(* CODESYS project EVs.export

Project tree, tasks and I/O mapping:
  visualisation EVs
*)

// /EVs
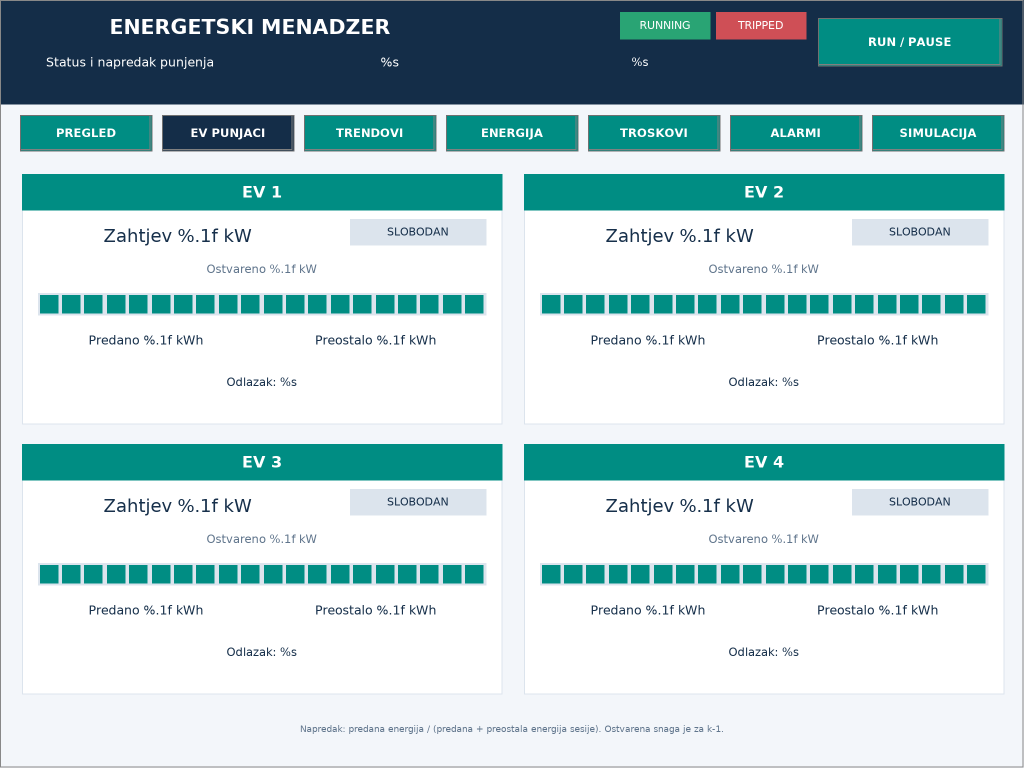
VISUALIZATION EVs  // 1024x768
    Rectangle (0,0 1024x768)
    Rectangle (0,0 1024x104)
    Rectangle (20,10 460x34), "ENERGETSKI MENADZER"
    Rectangle (20,48 220x28), "Status i napredak punjenja"
    Rectangle (260,49 260x26), "%s", text variable: Team_HMI.sDateTime
    Rectangle (530,49 220x26), "%s", text variable: Team_HMI.sPriceMode
    Button (818,18 184x48), "RUN / PAUSE"
        toggle SimCtrl.run
    Rectangle (620,12 90x27), "PAUSED", invisible if: SimCtrl.run
    Rectangle (620,12 90x27), "RUNNING", invisible if: NOT SimCtrl.run
    Rectangle (716,12 90x27), "TRIPPED", invisible if: NOT SimCtrl.tripped
    Button (20,115 132x36), "PREGLED"
        OnMouseClick:  Assign=Overview, Type=Assignment
    Button (162,115 132x36), "EV PUNJACI"
        OnMouseClick:  Assign=EVs, Type=Assignment
    Button (304,115 132x36), "TRENDOVI"
        OnMouseClick:  Assign=Trends, Type=Assignment
    Button (446,115 132x36), "ENERGIJA"
        OnMouseClick:  Assign=Energy, Type=Assignment
    Button (588,115 132x36), "TROSKOVI"
        OnMouseClick:  Assign=Costs, Type=Assignment
    Button (730,115 132x36), "ALARMI"
        OnMouseClick:  Assign=Alarms, Type=Assignment
    Button (872,115 132x36), "SIMULACIJA"
        OnMouseClick:  Assign=Controls, Type=Assignment
    Rectangle (22,174 480x250)
    Rectangle (22,174 480x36), "EV 1"
    Rectangle (350,219 136x26), "SPOJEN", invisible if: NOT Team_HMI.aEvConnected[0]
    Rectangle (350,219 136x26), "SLOBODAN", invisible if: Team_HMI.aEvConnected[0]
    Rectangle (38,218 280x36), "Zahtjev %.1f kW", text variable: Team_HMI.aEvReq[0]
    Rectangle (38,256 448x26), "Ostvareno %.1f kW", text variable: Team_HMI.aEvAct[0]
    Rectangle (38,293 448x22)
    Rectangle (40,295 18x18), invisible if: (100.0 * Team_HMI.aEvDelivered[0] / MAX(0.001, Team_HMI.aEvDelivered[0] + Team_HMI.aEvRemaining[0])) < 5.000
    Rectangle (62,295 18x18), invisible if: (100.0 * Team_HMI.aEvDelivered[0] / MAX(0.001, Team_HMI.aEvDelivered[0] + Team_HMI.aEvRemaining[0])) < 10.000
    Rectangle (84,295 18x18), invisible if: (100.0 * Team_HMI.aEvDelivered[0] / MAX(0.001, Team_HMI.aEvDelivered[0] + Team_HMI.aEvRemaining[0])) < 15.000
    Rectangle (107,295 18x18), invisible if: (100.0 * Team_HMI.aEvDelivered[0] / MAX(0.001, Team_HMI.aEvDelivered[0] + Team_HMI.aEvRemaining[0])) < 20.000
    Rectangle (129,295 18x18), invisible if: (100.0 * Team_HMI.aEvDelivered[0] / MAX(0.001, Team_HMI.aEvDelivered[0] + Team_HMI.aEvRemaining[0])) < 25.000
    Rectangle (152,295 18x18), invisible if: (100.0 * Team_HMI.aEvDelivered[0] / MAX(0.001, Team_HMI.aEvDelivered[0] + Team_HMI.aEvRemaining[0])) < 30.000
    Rectangle (174,295 18x18), invisible if: (100.0 * Team_HMI.aEvDelivered[0] / MAX(0.001, Team_HMI.aEvDelivered[0] + Team_HMI.aEvRemaining[0])) < 35.000
    Rectangle (196,295 18x18), invisible if: (100.0 * Team_HMI.aEvDelivered[0] / MAX(0.001, Team_HMI.aEvDelivered[0] + Team_HMI.aEvRemaining[0])) < 40.000
    Rectangle (219,295 18x18), invisible if: (100.0 * Team_HMI.aEvDelivered[0] / MAX(0.001, Team_HMI.aEvDelivered[0] + Team_HMI.aEvRemaining[0])) < 45.000
    Rectangle (241,295 18x18), invisible if: (100.0 * Team_HMI.aEvDelivered[0] / MAX(0.001, Team_HMI.aEvDelivered[0] + Team_HMI.aEvRemaining[0])) < 50.000
    Rectangle (264,295 18x18), invisible if: (100.0 * Team_HMI.aEvDelivered[0] / MAX(0.001, Team_HMI.aEvDelivered[0] + Team_HMI.aEvRemaining[0])) < 55.000
    Rectangle (286,295 18x18), invisible if: (100.0 * Team_HMI.aEvDelivered[0] / MAX(0.001, Team_HMI.aEvDelivered[0] + Team_HMI.aEvRemaining[0])) < 60.000
    Rectangle (308,295 18x18), invisible if: (100.0 * Team_HMI.aEvDelivered[0] / MAX(0.001, Team_HMI.aEvDelivered[0] + Team_HMI.aEvRemaining[0])) < 65.000
    Rectangle (331,295 18x18), invisible if: (100.0 * Team_HMI.aEvDelivered[0] / MAX(0.001, Team_HMI.aEvDelivered[0] + Team_HMI.aEvRemaining[0])) < 70.000
    Rectangle (353,295 18x18), invisible if: (100.0 * Team_HMI.aEvDelivered[0] / MAX(0.001, Team_HMI.aEvDelivered[0] + Team_HMI.aEvRemaining[0])) < 75.000
    Rectangle (376,295 18x18), invisible if: (100.0 * Team_HMI.aEvDelivered[0] / MAX(0.001, Team_HMI.aEvDelivered[0] + Team_HMI.aEvRemaining[0])) < 80.000
    Rectangle (398,295 18x18), invisible if: (100.0 * Team_HMI.aEvDelivered[0] / MAX(0.001, Team_HMI.aEvDelivered[0] + Team_HMI.aEvRemaining[0])) < 85.000
    Rectangle (420,295 18x18), invisible if: (100.0 * Team_HMI.aEvDelivered[0] / MAX(0.001, Team_HMI.aEvDelivered[0] + Team_HMI.aEvRemaining[0])) < 90.000
    Rectangle (443,295 18x18), invisible if: (100.0 * Team_HMI.aEvDelivered[0] / MAX(0.001, Team_HMI.aEvDelivered[0] + Team_HMI.aEvRemaining[0])) < 95.000
    Rectangle (465,295 18x18), invisible if: (100.0 * Team_HMI.aEvDelivered[0] / MAX(0.001, Team_HMI.aEvDelivered[0] + Team_HMI.aEvRemaining[0])) < 100.000
    Rectangle (38,325 216x30), "Predano %.1f kWh", text variable: Team_HMI.aEvDelivered[0]
    Rectangle (266,325 220x30), "Preostalo %.1f kWh", text variable: Team_HMI.aEvRemaining[0]
    Rectangle (38,367 448x30), "Odlazak: %s", text variable: Team_HMI.aEvDeparture[0]
    Rectangle (524,174 480x250)
    Rectangle (524,174 480x36), "EV 2"
    Rectangle (852,219 136x26), "SPOJEN", invisible if: NOT Team_HMI.aEvConnected[1]
    Rectangle (852,219 136x26), "SLOBODAN", invisible if: Team_HMI.aEvConnected[1]
    Rectangle (540,218 280x36), "Zahtjev %.1f kW", text variable: Team_HMI.aEvReq[1]
    Rectangle (540,256 448x26), "Ostvareno %.1f kW", text variable: Team_HMI.aEvAct[1]
    Rectangle (540,293 448x22)
    Rectangle (542,295 18x18), invisible if: (100.0 * Team_HMI.aEvDelivered[1] / MAX(0.001, Team_HMI.aEvDelivered[1] + Team_HMI.aEvRemaining[1])) < 5.000
    Rectangle (564,295 18x18), invisible if: (100.0 * Team_HMI.aEvDelivered[1] / MAX(0.001, Team_HMI.aEvDelivered[1] + Team_HMI.aEvRemaining[1])) < 10.000
    Rectangle (586,295 18x18), invisible if: (100.0 * Team_HMI.aEvDelivered[1] / MAX(0.001, Team_HMI.aEvDelivered[1] + Team_HMI.aEvRemaining[1])) < 15.000
    Rectangle (609,295 18x18), invisible if: (100.0 * Team_HMI.aEvDelivered[1] / MAX(0.001, Team_HMI.aEvDelivered[1] + Team_HMI.aEvRemaining[1])) < 20.000
    Rectangle (631,295 18x18), invisible if: (100.0 * Team_HMI.aEvDelivered[1] / MAX(0.001, Team_HMI.aEvDelivered[1] + Team_HMI.aEvRemaining[1])) < 25.000
    Rectangle (654,295 18x18), invisible if: (100.0 * Team_HMI.aEvDelivered[1] / MAX(0.001, Team_HMI.aEvDelivered[1] + Team_HMI.aEvRemaining[1])) < 30.000
    Rectangle (676,295 18x18), invisible if: (100.0 * Team_HMI.aEvDelivered[1] / MAX(0.001, Team_HMI.aEvDelivered[1] + Team_HMI.aEvRemaining[1])) < 35.000
    Rectangle (698,295 18x18), invisible if: (100.0 * Team_HMI.aEvDelivered[1] / MAX(0.001, Team_HMI.aEvDelivered[1] + Team_HMI.aEvRemaining[1])) < 40.000
    Rectangle (721,295 18x18), invisible if: (100.0 * Team_HMI.aEvDelivered[1] / MAX(0.001, Team_HMI.aEvDelivered[1] + Team_HMI.aEvRemaining[1])) < 45.000
    Rectangle (743,295 18x18), invisible if: (100.0 * Team_HMI.aEvDelivered[1] / MAX(0.001, Team_HMI.aEvDelivered[1] + Team_HMI.aEvRemaining[1])) < 50.000
    Rectangle (766,295 18x18), invisible if: (100.0 * Team_HMI.aEvDelivered[1] / MAX(0.001, Team_HMI.aEvDelivered[1] + Team_HMI.aEvRemaining[1])) < 55.000
    Rectangle (788,295 18x18), invisible if: (100.0 * Team_HMI.aEvDelivered[1] / MAX(0.001, Team_HMI.aEvDelivered[1] + Team_HMI.aEvRemaining[1])) < 60.000
    Rectangle (810,295 18x18), invisible if: (100.0 * Team_HMI.aEvDelivered[1] / MAX(0.001, Team_HMI.aEvDelivered[1] + Team_HMI.aEvRemaining[1])) < 65.000
    Rectangle (833,295 18x18), invisible if: (100.0 * Team_HMI.aEvDelivered[1] / MAX(0.001, Team_HMI.aEvDelivered[1] + Team_HMI.aEvRemaining[1])) < 70.000
    Rectangle (855,295 18x18), invisible if: (100.0 * Team_HMI.aEvDelivered[1] / MAX(0.001, Team_HMI.aEvDelivered[1] + Team_HMI.aEvRemaining[1])) < 75.000
    Rectangle (878,295 18x18), invisible if: (100.0 * Team_HMI.aEvDelivered[1] / MAX(0.001, Team_HMI.aEvDelivered[1] + Team_HMI.aEvRemaining[1])) < 80.000
    Rectangle (900,295 18x18), invisible if: (100.0 * Team_HMI.aEvDelivered[1] / MAX(0.001, Team_HMI.aEvDelivered[1] + Team_HMI.aEvRemaining[1])) < 85.000
    Rectangle (922,295 18x18), invisible if: (100.0 * Team_HMI.aEvDelivered[1] / MAX(0.001, Team_HMI.aEvDelivered[1] + Team_HMI.aEvRemaining[1])) < 90.000
    Rectangle (945,295 18x18), invisible if: (100.0 * Team_HMI.aEvDelivered[1] / MAX(0.001, Team_HMI.aEvDelivered[1] + Team_HMI.aEvRemaining[1])) < 95.000
    Rectangle (967,295 18x18), invisible if: (100.0 * Team_HMI.aEvDelivered[1] / MAX(0.001, Team_HMI.aEvDelivered[1] + Team_HMI.aEvRemaining[1])) < 100.000
    Rectangle (540,325 216x30), "Predano %.1f kWh", text variable: Team_HMI.aEvDelivered[1]
    Rectangle (768,325 220x30), "Preostalo %.1f kWh", text variable: Team_HMI.aEvRemaining[1]
    Rectangle (540,367 448x30), "Odlazak: %s", text variable: Team_HMI.aEvDeparture[1]
    Rectangle (22,444 480x250)
    Rectangle (22,444 480x36), "EV 3"
    Rectangle (350,489 136x26), "SPOJEN", invisible if: NOT Team_HMI.aEvConnected[2]
    Rectangle (350,489 136x26), "SLOBODAN", invisible if: Team_HMI.aEvConnected[2]
    Rectangle (38,488 280x36), "Zahtjev %.1f kW", text variable: Team_HMI.aEvReq[2]
    Rectangle (38,526 448x26), "Ostvareno %.1f kW", text variable: Team_HMI.aEvAct[2]
    Rectangle (38,563 448x22)
    Rectangle (40,565 18x18), invisible if: (100.0 * Team_HMI.aEvDelivered[2] / MAX(0.001, Team_HMI.aEvDelivered[2] + Team_HMI.aEvRemaining[2])) < 5.000
    Rectangle (62,565 18x18), invisible if: (100.0 * Team_HMI.aEvDelivered[2] / MAX(0.001, Team_HMI.aEvDelivered[2] + Team_HMI.aEvRemaining[2])) < 10.000
    Rectangle (84,565 18x18), invisible if: (100.0 * Team_HMI.aEvDelivered[2] / MAX(0.001, Team_HMI.aEvDelivered[2] + Team_HMI.aEvRemaining[2])) < 15.000
    Rectangle (107,565 18x18), invisible if: (100.0 * Team_HMI.aEvDelivered[2] / MAX(0.001, Team_HMI.aEvDelivered[2] + Team_HMI.aEvRemaining[2])) < 20.000
    Rectangle (129,565 18x18), invisible if: (100.0 * Team_HMI.aEvDelivered[2] / MAX(0.001, Team_HMI.aEvDelivered[2] + Team_HMI.aEvRemaining[2])) < 25.000
    Rectangle (152,565 18x18), invisible if: (100.0 * Team_HMI.aEvDelivered[2] / MAX(0.001, Team_HMI.aEvDelivered[2] + Team_HMI.aEvRemaining[2])) < 30.000
    Rectangle (174,565 18x18), invisible if: (100.0 * Team_HMI.aEvDelivered[2] / MAX(0.001, Team_HMI.aEvDelivered[2] + Team_HMI.aEvRemaining[2])) < 35.000
    Rectangle (196,565 18x18), invisible if: (100.0 * Team_HMI.aEvDelivered[2] / MAX(0.001, Team_HMI.aEvDelivered[2] + Team_HMI.aEvRemaining[2])) < 40.000
    Rectangle (219,565 18x18), invisible if: (100.0 * Team_HMI.aEvDelivered[2] / MAX(0.001, Team_HMI.aEvDelivered[2] + Team_HMI.aEvRemaining[2])) < 45.000
    Rectangle (241,565 18x18), invisible if: (100.0 * Team_HMI.aEvDelivered[2] / MAX(0.001, Team_HMI.aEvDelivered[2] + Team_HMI.aEvRemaining[2])) < 50.000
    Rectangle (264,565 18x18), invisible if: (100.0 * Team_HMI.aEvDelivered[2] / MAX(0.001, Team_HMI.aEvDelivered[2] + Team_HMI.aEvRemaining[2])) < 55.000
    Rectangle (286,565 18x18), invisible if: (100.0 * Team_HMI.aEvDelivered[2] / MAX(0.001, Team_HMI.aEvDelivered[2] + Team_HMI.aEvRemaining[2])) < 60.000
    Rectangle (308,565 18x18), invisible if: (100.0 * Team_HMI.aEvDelivered[2] / MAX(0.001, Team_HMI.aEvDelivered[2] + Team_HMI.aEvRemaining[2])) < 65.000
    Rectangle (331,565 18x18), invisible if: (100.0 * Team_HMI.aEvDelivered[2] / MAX(0.001, Team_HMI.aEvDelivered[2] + Team_HMI.aEvRemaining[2])) < 70.000
    Rectangle (353,565 18x18), invisible if: (100.0 * Team_HMI.aEvDelivered[2] / MAX(0.001, Team_HMI.aEvDelivered[2] + Team_HMI.aEvRemaining[2])) < 75.000
    Rectangle (376,565 18x18), invisible if: (100.0 * Team_HMI.aEvDelivered[2] / MAX(0.001, Team_HMI.aEvDelivered[2] + Team_HMI.aEvRemaining[2])) < 80.000
    Rectangle (398,565 18x18), invisible if: (100.0 * Team_HMI.aEvDelivered[2] / MAX(0.001, Team_HMI.aEvDelivered[2] + Team_HMI.aEvRemaining[2])) < 85.000
    Rectangle (420,565 18x18), invisible if: (100.0 * Team_HMI.aEvDelivered[2] / MAX(0.001, Team_HMI.aEvDelivered[2] + Team_HMI.aEvRemaining[2])) < 90.000
    Rectangle (443,565 18x18), invisible if: (100.0 * Team_HMI.aEvDelivered[2] / MAX(0.001, Team_HMI.aEvDelivered[2] + Team_HMI.aEvRemaining[2])) < 95.000
    Rectangle (465,565 18x18), invisible if: (100.0 * Team_HMI.aEvDelivered[2] / MAX(0.001, Team_HMI.aEvDelivered[2] + Team_HMI.aEvRemaining[2])) < 100.000
    Rectangle (38,595 216x30), "Predano %.1f kWh", text variable: Team_HMI.aEvDelivered[2]
    Rectangle (266,595 220x30), "Preostalo %.1f kWh", text variable: Team_HMI.aEvRemaining[2]
    Rectangle (38,637 448x30), "Odlazak: %s", text variable: Team_HMI.aEvDeparture[2]
    Rectangle (524,444 480x250)
    Rectangle (524,444 480x36), "EV 4"
    Rectangle (852,489 136x26), "SPOJEN", invisible if: NOT Team_HMI.aEvConnected[3]
    Rectangle (852,489 136x26), "SLOBODAN", invisible if: Team_HMI.aEvConnected[3]
    Rectangle (540,488 280x36), "Zahtjev %.1f kW", text variable: Team_HMI.aEvReq[3]
    Rectangle (540,526 448x26), "Ostvareno %.1f kW", text variable: Team_HMI.aEvAct[3]
    Rectangle (540,563 448x22)
    Rectangle (542,565 18x18), invisible if: (100.0 * Team_HMI.aEvDelivered[3] / MAX(0.001, Team_HMI.aEvDelivered[3] + Team_HMI.aEvRemaining[3])) < 5.000
    Rectangle (564,565 18x18), invisible if: (100.0 * Team_HMI.aEvDelivered[3] / MAX(0.001, Team_HMI.aEvDelivered[3] + Team_HMI.aEvRemaining[3])) < 10.000
    Rectangle (586,565 18x18), invisible if: (100.0 * Team_HMI.aEvDelivered[3] / MAX(0.001, Team_HMI.aEvDelivered[3] + Team_HMI.aEvRemaining[3])) < 15.000
    Rectangle (609,565 18x18), invisible if: (100.0 * Team_HMI.aEvDelivered[3] / MAX(0.001, Team_HMI.aEvDelivered[3] + Team_HMI.aEvRemaining[3])) < 20.000
    Rectangle (631,565 18x18), invisible if: (100.0 * Team_HMI.aEvDelivered[3] / MAX(0.001, Team_HMI.aEvDelivered[3] + Team_HMI.aEvRemaining[3])) < 25.000
    Rectangle (654,565 18x18), invisible if: (100.0 * Team_HMI.aEvDelivered[3] / MAX(0.001, Team_HMI.aEvDelivered[3] + Team_HMI.aEvRemaining[3])) < 30.000
    Rectangle (676,565 18x18), invisible if: (100.0 * Team_HMI.aEvDelivered[3] / MAX(0.001, Team_HMI.aEvDelivered[3] + Team_HMI.aEvRemaining[3])) < 35.000
    Rectangle (698,565 18x18), invisible if: (100.0 * Team_HMI.aEvDelivered[3] / MAX(0.001, Team_HMI.aEvDelivered[3] + Team_HMI.aEvRemaining[3])) < 40.000
    Rectangle (721,565 18x18), invisible if: (100.0 * Team_HMI.aEvDelivered[3] / MAX(0.001, Team_HMI.aEvDelivered[3] + Team_HMI.aEvRemaining[3])) < 45.000
    Rectangle (743,565 18x18), invisible if: (100.0 * Team_HMI.aEvDelivered[3] / MAX(0.001, Team_HMI.aEvDelivered[3] + Team_HMI.aEvRemaining[3])) < 50.000
    Rectangle (766,565 18x18), invisible if: (100.0 * Team_HMI.aEvDelivered[3] / MAX(0.001, Team_HMI.aEvDelivered[3] + Team_HMI.aEvRemaining[3])) < 55.000
    Rectangle (788,565 18x18), invisible if: (100.0 * Team_HMI.aEvDelivered[3] / MAX(0.001, Team_HMI.aEvDelivered[3] + Team_HMI.aEvRemaining[3])) < 60.000
    Rectangle (810,565 18x18), invisible if: (100.0 * Team_HMI.aEvDelivered[3] / MAX(0.001, Team_HMI.aEvDelivered[3] + Team_HMI.aEvRemaining[3])) < 65.000
    Rectangle (833,565 18x18), invisible if: (100.0 * Team_HMI.aEvDelivered[3] / MAX(0.001, Team_HMI.aEvDelivered[3] + Team_HMI.aEvRemaining[3])) < 70.000
    Rectangle (855,565 18x18), invisible if: (100.0 * Team_HMI.aEvDelivered[3] / MAX(0.001, Team_HMI.aEvDelivered[3] + Team_HMI.aEvRemaining[3])) < 75.000
    Rectangle (878,565 18x18), invisible if: (100.0 * Team_HMI.aEvDelivered[3] / MAX(0.001, Team_HMI.aEvDelivered[3] + Team_HMI.aEvRemaining[3])) < 80.000
    Rectangle (900,565 18x18), invisible if: (100.0 * Team_HMI.aEvDelivered[3] / MAX(0.001, Team_HMI.aEvDelivered[3] + Team_HMI.aEvRemaining[3])) < 85.000
    Rectangle (922,565 18x18), invisible if: (100.0 * Team_HMI.aEvDelivered[3] / MAX(0.001, Team_HMI.aEvDelivered[3] + Team_HMI.aEvRemaining[3])) < 90.000
    Rectangle (945,565 18x18), invisible if: (100.0 * Team_HMI.aEvDelivered[3] / MAX(0.001, Team_HMI.aEvDelivered[3] + Team_HMI.aEvRemaining[3])) < 95.000
    Rectangle (967,565 18x18), invisible if: (100.0 * Team_HMI.aEvDelivered[3] / MAX(0.001, Team_HMI.aEvDelivered[3] + Team_HMI.aEvRemaining[3])) < 100.000
    Rectangle (540,595 216x30), "Predano %.1f kWh", text variable: Team_HMI.aEvDelivered[3]
    Rectangle (768,595 220x30), "Preostalo %.1f kWh", text variable: Team_HMI.aEvRemaining[3]
    Rectangle (540,637 448x30), "Odlazak: %s", text variable: Team_HMI.aEvDeparture[3]
    Rectangle (22,718 980x22), "Napredak: predana energija / (predana + preostala energija sesije). Ostvarena snaga je za k-1."
END_VISUALIZATION
